(* IEC 61131-3 sources: rusty/tests/lit/single/type_promotion/bit_string/comparison, 10 files *)

(* ---- byte_word_variables.st ---- *)
// RUN: %COMPILE %s && %RUN | %CHECK %s
// Two BYTE or WORD operands keep their own width and compare unsigned, so a value from the signed midpoint on compares as large.
FUNCTION main : DINT
    VAR
        bhi : BYTE := 16#FF;
        blo : BYTE := 16#01;
        bmid : BYTE := 16#80;
        bbelow : BYTE := 16#7F;
        whi : WORD := 16#FFFF;
        wlo : WORD := 16#0001;
        wmid : WORD := 16#8000;
        wbelow : WORD := 16#7FFF;
    END_VAR

    // BYTE
    printf('BYTE hi > lo = %d$N', bhi > blo);               // CHECK: BYTE hi > lo = 1
    printf('BYTE lo < hi = %d$N', blo < bhi);               // CHECK-NEXT: BYTE lo < hi = 1
    printf('BYTE hi <= lo = %d$N', bhi <= blo);             // CHECK-NEXT: BYTE hi <= lo = 0
    printf('BYTE mid > below = %d$N', bmid > bbelow);       // CHECK-NEXT: BYTE mid > below = 1
    printf('BYTE hi > BYTE#1 = %d$N', bhi > BYTE#1);        // CHECK-NEXT: BYTE hi > BYTE#1 = 1

    // WORD
    printf('WORD hi > lo = %d$N', whi > wlo);               // CHECK-NEXT: WORD hi > lo = 1
    printf('WORD lo < hi = %d$N', wlo < whi);               // CHECK-NEXT: WORD lo < hi = 1
    printf('WORD hi <= lo = %d$N', whi <= wlo);             // CHECK-NEXT: WORD hi <= lo = 0
    printf('WORD mid > below = %d$N', wmid > wbelow);       // CHECK-NEXT: WORD mid > below = 1
    printf('WORD hi > WORD#1 = %d$N', whi > WORD#1);        // CHECK-NEXT: WORD hi > WORD#1 = 1
END_FUNCTION

(* ---- compare_guards.st ---- *)
// RUN: %COMPILE %s && %RUN | %CHECK %s
// Bit string compares whose result does not depend on the signedness of the predicate.
FUNCTION main : DINT
    VAR
        dw : DWORD := 16#FFFF_FFFF;
        lw : LWORD := 16#FFFF_FFFF_FFFF_FFFF;
        b : BYTE := 16#FF;
        w : WORD := 16#FFFF;
        im1 : INT := -1;
    END_VAR

    // Equality compares the bit pattern
    printf('DWORD 16#FFFF_FFFF = -1 = %d$N', dw = -1);      // CHECK: DWORD 16#FFFF_FFFF = -1 = 1
    printf('LWORD max = 16#FFFF_FFFF_FFFF_FFFF = %d$N', lw = 16#FFFF_FFFF_FFFF_FFFF);    // CHECK-NEXT: LWORD max = 16#FFFF_FFFF_FFFF_FFFF = 1

    // A narrow bit string next to an untyped literal is widened to DINT
    printf('BYTE 16#FF > 1 = %d$N', b > 1);                 // CHECK-NEXT: BYTE 16#FF > 1 = 1
    printf('WORD 16#FFFF > 1 = %d$N', w > 1);               // CHECK-NEXT: WORD 16#FFFF > 1 = 1

    // Results that hold under either predicate
    printf('INT -1 > DWORD max = %d$N', im1 > dw);          // CHECK-NEXT: INT -1 > DWORD max = 0
END_FUNCTION

(* ---- dword_variables.st ---- *)
// RUN: %COMPILE %s && %RUN | %CHECK %s
// A relational compare of two DWORD values is unsigned, so a value from the signed midpoint on compares as large.
FUNCTION main : DINT
    VAR
        hi : DWORD := 16#FFFF_FFFF;
        lo : DWORD := 16#1;
        mid : DWORD := 16#8000_0000;
        below : DWORD := 16#7FFF_FFFF;
        result : BOOL;
    END_VAR

    // Every relational operator, both operand orders
    printf('hi > lo = %d$N', hi > lo);             // CHECK: hi > lo = 1
    printf('hi >= lo = %d$N', hi >= lo);           // CHECK-NEXT: hi >= lo = 1
    printf('hi < lo = %d$N', hi < lo);             // CHECK-NEXT: hi < lo = 0
    printf('hi <= lo = %d$N', hi <= lo);           // CHECK-NEXT: hi <= lo = 0
    printf('lo < hi = %d$N', lo < hi);             // CHECK-NEXT: lo < hi = 1
    printf('lo <= hi = %d$N', lo <= hi);           // CHECK-NEXT: lo <= hi = 1
    printf('lo > hi = %d$N', lo > hi);             // CHECK-NEXT: lo > hi = 0
    printf('lo >= hi = %d$N', lo >= hi);           // CHECK-NEXT: lo >= hi = 0

    // The two values next to the signed midpoint
    printf('mid > below = %d$N', mid > below);     // CHECK-NEXT: mid > below = 1

    // A typed literal operand of the same type
    printf('hi > DWORD#16#1 = %d$N', hi > DWORD#16#1);  // CHECK-NEXT: hi > DWORD#16#1 = 1

    // The compare as a stored value and as a condition
    result := hi > lo;
    printf('stored = %d$N', result);               // CHECK-NEXT: stored = 1
    IF hi > lo THEN
        printf('IF taken$N');                      // CHECK-NEXT: IF taken
    ELSE
        printf('IF not taken$N');
    END_IF
END_FUNCTION

(* ---- lword_variables.st ---- *)
// RUN: %COMPILE %s && %RUN | %CHECK %s
// A relational compare of two LWORD values is unsigned, so a value from the signed midpoint on compares as large.
FUNCTION main : DINT
    VAR
        hi : LWORD := 16#FFFF_FFFF_FFFF_FFFF;
        lo : LWORD := 16#1;
        mid : LWORD := 16#8000_0000_0000_0000;
        below : LWORD := 16#7FFF_FFFF_FFFF_FFFF;
        result : BOOL;
    END_VAR

    // Every relational operator, both operand orders
    printf('hi > lo = %d$N', hi > lo);             // CHECK: hi > lo = 1
    printf('hi >= lo = %d$N', hi >= lo);           // CHECK-NEXT: hi >= lo = 1
    printf('hi < lo = %d$N', hi < lo);             // CHECK-NEXT: hi < lo = 0
    printf('hi <= lo = %d$N', hi <= lo);           // CHECK-NEXT: hi <= lo = 0
    printf('lo < hi = %d$N', lo < hi);             // CHECK-NEXT: lo < hi = 1
    printf('lo <= hi = %d$N', lo <= hi);           // CHECK-NEXT: lo <= hi = 1
    printf('lo > hi = %d$N', lo > hi);             // CHECK-NEXT: lo > hi = 0
    printf('lo >= hi = %d$N', lo >= hi);           // CHECK-NEXT: lo >= hi = 0

    // The two values next to the signed midpoint
    printf('mid > below = %d$N', mid > below);     // CHECK-NEXT: mid > below = 1

    // A typed literal operand of the same type
    printf('hi > LWORD#16#1 = %d$N', hi > LWORD#16#1);  // CHECK-NEXT: hi > LWORD#16#1 = 1

    // The compare as a stored value and as a condition
    result := hi > lo;
    printf('stored = %d$N', result);               // CHECK-NEXT: stored = 1
    IF hi > lo THEN
        printf('IF taken$N');                      // CHECK-NEXT: IF taken
    ELSE
        printf('IF not taken$N');
    END_IF
END_FUNCTION

(* ---- mixed_width_bit_strings.st ---- *)
// RUN: %COMPILE %s && %RUN | %CHECK %s
// A BYTE and a WORD operand keep the wider bit string type and compare unsigned, so a value from the signed midpoint on compares as large.
FUNCTION main : DINT
    VAR
        b5 : BYTE := 16#05;
        b2 : BYTE := 16#02;
        wmax : WORD := 16#FFFF;
    END_VAR

    printf('BYTE 5 < WORD max = %d$N', b5 < wmax);          // CHECK: BYTE 5 < WORD max = 1
    printf('BYTE 5 > WORD max = %d$N', b5 > wmax);          // CHECK-NEXT: BYTE 5 > WORD max = 0
    printf('WORD max > BYTE 2 = %d$N', wmax > b2);          // CHECK-NEXT: WORD max > BYTE 2 = 1
    printf('WORD max < BYTE 2 = %d$N', wmax < b2);          // CHECK-NEXT: WORD max < BYTE 2 = 0
END_FUNCTION

(* ---- mixed_width_with_unsigned_integers.st ---- *)
// RUN: %COMPILE %s && %RUN | %CHECK %s
// A bit string next to an unsigned integer or another bit string of a different width is promoted to the wider 32-bit or 64-bit type
// and then compared unsigned.
FUNCTION main : DINT
    VAR
        us5 : USINT := 5;
        ui5 : UINT := 5;
        b5 : BYTE := 16#05;
        w5 : WORD := 16#0005;
        ud5 : UDINT := 5;
        dw5 : DWORD := 16#5;
        us2 : USINT := 2;
        ui2 : UINT := 2;
        ud2 : UDINT := 2;
        dw2 : DWORD := 16#2;
        lw2 : LWORD := 16#2;
        udmax : UDINT := 4294967295;
        dwmax : DWORD := 16#FFFF_FFFF;
        ulmax : ULINT := 18446744073709551615;
        lwmax : LWORD := 16#FFFF_FFFF_FFFF_FFFF;
    END_VAR

    // Narrow operand next to a 32-bit maximum
    printf('UINT 5 < DWORD max = %d$N', ui5 < dwmax);       // CHECK: UINT 5 < DWORD max = 1
    printf('BYTE 5 < UDINT max = %d$N', b5 < udmax);        // CHECK-NEXT: BYTE 5 < UDINT max = 1
    printf('WORD 5 < DWORD max = %d$N', w5 < dwmax);        // CHECK-NEXT: WORD 5 < DWORD max = 1
    printf('DWORD max > UINT 2 = %d$N', dwmax > ui2);       // CHECK-NEXT: DWORD max > UINT 2 = 1

    // Narrow operand next to a 64-bit maximum
    printf('BYTE 5 < LWORD max = %d$N', b5 < lwmax);        // CHECK-NEXT: BYTE 5 < LWORD max = 1
    printf('LWORD max > USINT 2 = %d$N', lwmax > us2);      // CHECK-NEXT: LWORD max > USINT 2 = 1

    // 32-bit operand next to a 64-bit maximum
    printf('DWORD 5 < LWORD max = %d$N', dw5 < lwmax);      // CHECK-NEXT: DWORD 5 < LWORD max = 1
    printf('UDINT 5 < LWORD max = %d$N', ud5 < lwmax);      // CHECK-NEXT: UDINT 5 < LWORD max = 1
    printf('ULINT max > DWORD 2 = %d$N', ulmax > dw2);      // CHECK-NEXT: ULINT max > DWORD 2 = 1
    printf('USINT 5 < DWORD max = %d$N', us5 < dwmax);      // CHECK-NEXT: USINT 5 < DWORD max = 1

    // Unsigned integer next to a bit string of the same width
    printf('UDINT max > DWORD 2 = %d$N', udmax > dw2);      // CHECK-NEXT: UDINT max > DWORD 2 = 1
    printf('DWORD max > UDINT 2 = %d$N', dwmax > ud2);      // CHECK-NEXT: DWORD max > UDINT 2 = 1
    printf('ULINT max > LWORD 2 = %d$N', ulmax > lw2);      // CHECK-NEXT: ULINT max > LWORD 2 = 1
END_FUNCTION

(* ---- with_negative_literal.st ---- *)
// RUN: %COMPILE %s && %RUN | %CHECK %s
// XFAIL: *
// A negative literal next to a DWORD or LWORD maximum compares signed, so the maximum reads as -1.
FUNCTION main : DINT
    VAR
        dwmax : DWORD := 16#FFFF_FFFF;
        lwmax : LWORD := 16#FFFF_FFFF_FFFF_FFFF;
    END_VAR

    printf('DWORD max > -1 = %d$N', dwmax > -1);            // CHECK: DWORD max > -1 = 1
    printf('LWORD max > -1 = %d$N', lwmax > -1);            // CHECK-NEXT: LWORD max > -1 = 1
    printf('-1 < DWORD max = %d$N', -1 < dwmax);            // CHECK-NEXT: -1 < DWORD max = 1
END_FUNCTION

(* ---- with_signed_operand.st ---- *)
// RUN: %COMPILE %s && %RUN | %CHECK %s
// XFAIL: *
// A signed operand next to a DWORD or LWORD makes the compare signed, so a bit string from the signed midpoint on compares as negative.
FUNCTION main : DINT
    VAR
        i5 : INT := 5;
        im1 : INT := -1;
        dm1 : DINT := -1;
        lm1 : LINT := -1;
        i2 : INT := 2;
        l2 : LINT := 2;
        dwmax : DWORD := 16#FFFF_FFFF;
        lwmax : LWORD := 16#FFFF_FFFF_FFFF_FFFF;
    END_VAR

    // Signed value below a bit string maximum
    printf('INT 5 < DWORD max = %d$N', i5 < dwmax);         // CHECK: INT 5 < DWORD max = 1
    printf('INT -1 < DWORD max = %d$N', im1 < dwmax);       // CHECK-NEXT: INT -1 < DWORD max = 1
    printf('LINT -1 < LWORD max = %d$N', lm1 < lwmax);      // CHECK-NEXT: LINT -1 < LWORD max = 1

    // Bit string maximum on the left
    printf('DWORD max > INT 2 = %d$N', dwmax > i2);         // CHECK-NEXT: DWORD max > INT 2 = 1
    printf('LWORD max > DINT -1 = %d$N', lwmax > dm1);      // CHECK-NEXT: LWORD max > DINT -1 = 1
    printf('LWORD max > LINT 2 = %d$N', lwmax > l2);        // CHECK-NEXT: LWORD max > LINT 2 = 1
END_FUNCTION

(* ---- with_untyped_literal.st ---- *)
// RUN: %COMPILE %s && %RUN | %CHECK %s
// An untyped integer literal takes the type of a DWORD or LWORD operand, so the compare is unsigned.
FUNCTION main : DINT
    VAR
        dw : DWORD := 16#FFFF_FFFF;
        lw : LWORD := 16#FFFF_FFFF_FFFF_FFFF;
    END_VAR

    // Literal on the right
    printf('DWORD > 1 = %d$N', dw > 1);                     // CHECK: DWORD > 1 = 1
    printf('DWORD > 16#7FFF_FFFF = %d$N', dw > 16#7FFF_FFFF);   // CHECK-NEXT: DWORD > 16#7FFF_FFFF = 1
    printf('DWORD < 0 = %d$N', dw < 0);                     // CHECK-NEXT: DWORD < 0 = 0
    printf('LWORD > 1 = %d$N', lw > 1);                     // CHECK-NEXT: LWORD > 1 = 1
    printf('LWORD > 3000000000 = %d$N', lw > 3000000000);   // CHECK-NEXT: LWORD > 3000000000 = 1

    // Literal on the left
    printf('1 < DWORD = %d$N', 1 < dw);                     // CHECK-NEXT: 1 < DWORD = 1
    printf('1 < LWORD = %d$N', 1 < lw);                     // CHECK-NEXT: 1 < LWORD = 1
END_FUNCTION

(* ---- literal_by_declaration_section.st ---- *)
// RUN: %COMPILE %s && %RUN | %CHECK %s
// A compare of a DWORD or LWORD operand with an untyped literal is unsigned, wherever the operand is declared.
VAR_GLOBAL
    g : DWORD := 16#FFFF_FFFF;
END_VAR

VAR_GLOBAL CONSTANT
    gc : LWORD := 16#FFFF_FFFF_FFFF_FFFF;
END_VAR

FUNCTION_BLOCK probe
    VAR_INPUT
        i : DWORD;
    END_VAR
    VAR_INPUT CONSTANT
        ic : DWORD := 16#FFFF_FFFF;
    END_VAR
    VAR_IN_OUT
        io : LWORD;
    END_VAR
    VAR_OUTPUT
        o : DWORD;
    END_VAR
    VAR
        m : LWORD := 16#FFFF_FFFF_FFFF_FFFF;
    END_VAR
    VAR CONSTANT
        c : DWORD := 16#FFFF_FFFF;
    END_VAR
    VAR_TEMP
        t : DWORD;
    END_VAR

    o := 16#FFFF_FFFF;
    t := 16#FFFF_FFFF;
    printf('VAR_INPUT > 16#7FFFFFFF = %d$N', i > 16#7FFFFFFF);
    printf('VAR_INPUT CONSTANT < 0 = %d$N', ic < 0);
    printf('VAR_IN_OUT > 16#7FFFFFFF = %d$N', io > 16#7FFFFFFF);
    printf('VAR_OUTPUT < 0 = %d$N', o < 0);
    printf('VAR > 3000000000 = %d$N', m > 3000000000);
    printf('VAR CONSTANT > 16#7FFFFFFF = %d$N', c > 16#7FFFFFFF);
    printf('VAR_TEMP < 0 = %d$N', t < 0);
    printf('VAR_GLOBAL > 16#7FFFFFFF = %d$N', g > 16#7FFFFFFF);
    printf('VAR_GLOBAL CONSTANT < 0 = %d$N', gc < 0);
END_FUNCTION_BLOCK

FUNCTION main : DINT
    VAR
        inst : probe;
        v : LWORD := 16#FFFF_FFFF_FFFF_FFFF;
    END_VAR

    inst(i := 16#FFFF_FFFF, io := v);
    // CHECK: VAR_INPUT > 16#7FFFFFFF = 1
    // CHECK-NEXT: VAR_INPUT CONSTANT < 0 = 0
    // CHECK-NEXT: VAR_IN_OUT > 16#7FFFFFFF = 1
    // CHECK-NEXT: VAR_OUTPUT < 0 = 0
    // CHECK-NEXT: VAR > 3000000000 = 1
    // CHECK-NEXT: VAR CONSTANT > 16#7FFFFFFF = 1
    // CHECK-NEXT: VAR_TEMP < 0 = 0
    // CHECK-NEXT: VAR_GLOBAL > 16#7FFFFFFF = 1
    // CHECK-NEXT: VAR_GLOBAL CONSTANT < 0 = 0
END_FUNCTION
